TYPE stShutterCmdEvent :
STRUCT
	Execute : BOOL;
    Cmd : stShutterCmd;
	Source  : eShutterCmdSource;
END_STRUCT
END_TYPE

(* stored: Version 1.1.0.1
   DUT stShutterCmdEvent: Id {e6ee52d5-e2da-4fe0-b612-a98cede1bba8} *)
